INTERFACE I_LintItf

METHOD M_Do : BOOL
VAR_INPUT
END_VAR
END_METHOD

PROPERTY P_Val : INT
END_PROPERTY

END_INTERFACE

(* stored: Version 1.1.0.1, ProductVersion 3.1.4024.16
   Itf I_LintItf: Id {9d0ff248-6f43-44db-b865-b80230e2ba0a}
   Method M_Do: Id {13aa9473-a3ca-476a-b49e-2680cb04806e}
   Property P_Val: Id {8a4b6363-03be-49da-a4df-2f05238b4419} *)
